PROGRAM PRG_Seq
VAR
    eStep, ePrevStep : E_Step := E_Step.eInit;
    nFaultCode       : UINT;        // 1=E-stop 2=no air 3=cylinder fault 4=step timeout
    nPartCount       : UDINT;
    bRejectPart      : BOOL;
    xAutoRun         : BOOL;
    xReady           : BOOL;
    xEnableCyl       : BOOL;

    // cylinder commands (TRUE = working position AS, FALSE = home GS) - persistent
    xInfeedWork, xClampWork, xEjectWork, xDivertWork, xOutfeedWork : BOOL;
    // momentary commands (cleared every scan, set by the active step)
    xBlow, xBypass, xLaserOn, xTrig : BOOL;

    fbInfeed, fbOutfeed, fbEjector, fbClamp, fbDiverter : FB_Cylinder;
    rStart, rReset   : R_TRIG;
    fbPart           : TON;
    fbBlowTime       : TON;
    fbStepTO         : TON;
    tStepTimeout     : TIME := T#30S;
    tBlow            : TIME := T#1S;
    tPartDebounce    : TIME := T#200MS;
END_VAR

rStart(CLK := GVL_Ctrl.xStart);
rReset(CLK := GVL_Ctrl.xReset);
IF rStart.Q THEN xAutoRun := TRUE;  END_IF
IF GVL_Ctrl.xStop THEN xAutoRun := FALSE; END_IF

// momentary outputs default to OFF every scan
xBlow := FALSE;  xBypass := FALSE;  xLaserOn := FALSE;  xTrig := FALSE;

xReady := GVL_IO.xPressureOK AND NOT GVL_IO.xEStop
          AND GVL_IO.xServoInLatched AND GVL_IO.xServoOutLatched;
xEnableCyl := (eStep <> E_Step.eFault) AND NOT GVL_IO.xEStop AND GVL_IO.xPressureOK;

// ---- cylinders (called first so that feedback is current for the transitions)
fbInfeed(  xCmdWork := xInfeedWork,  xEnable := xEnableCyl, xReset := rReset.Q,
           xSensWork := GVL_IO.stInfeed.xSensWork,   xSensHome := GVL_IO.stInfeed.xSensHome,
           xValveWork => GVL_IO.stInfeed.xValveWork, xValveHome => GVL_IO.stInfeed.xValveHome);
fbOutfeed( xCmdWork := xOutfeedWork, xEnable := xEnableCyl, xReset := rReset.Q,
           xSensWork := GVL_IO.stOutfeed.xSensWork,   xSensHome := GVL_IO.stOutfeed.xSensHome,
           xValveWork => GVL_IO.stOutfeed.xValveWork, xValveHome => GVL_IO.stOutfeed.xValveHome);
fbEjector( xCmdWork := xEjectWork,   xEnable := xEnableCyl, xReset := rReset.Q,
           xSensWork := GVL_IO.stEjector.xSensWork,   xSensHome := GVL_IO.stEjector.xSensHome,
           xValveWork => GVL_IO.stEjector.xValveWork, xValveHome => GVL_IO.stEjector.xValveHome);
fbClamp(   xCmdWork := xClampWork,   xEnable := xEnableCyl, xReset := rReset.Q,
           xSensWork := GVL_IO.stClamp.xSensWork,   xSensHome := GVL_IO.stClamp.xSensHome,
           xValveWork => GVL_IO.stClamp.xValveWork, xValveHome => GVL_IO.stClamp.xValveHome);
fbDiverter(xCmdWork := xDivertWork,  xEnable := xEnableCyl, xReset := rReset.Q,
           xSensWork := GVL_IO.stDiverter.xSensWork,   xSensHome := GVL_IO.stDiverter.xSensHome,
           xValveWork => GVL_IO.stDiverter.xValveWork, xValveHome => GVL_IO.stDiverter.xValveHome);

// ---- step timeout (restarts whenever the step changes)
fbStepTO(IN := (eStep = ePrevStep) AND (eStep <> E_Step.eIdle) AND (eStep <> E_Step.eWaitPart)
               AND (eStep <> E_Step.eFault),
         PT := tStepTimeout);
ePrevStep := eStep;

// ---- supervision
IF eStep <> E_Step.eFault THEN
    IF GVL_IO.xEStop THEN
        nFaultCode := 1;  eStep := E_Step.eFault;
    ELSIF NOT GVL_IO.xPressureOK THEN
        nFaultCode := 2;  eStep := E_Step.eFault;
    ELSIF fbInfeed.xFault OR fbOutfeed.xFault OR fbEjector.xFault OR fbClamp.xFault OR fbDiverter.xFault THEN
        nFaultCode := 3;  eStep := E_Step.eFault;
    ELSIF fbStepTO.Q THEN
        nFaultCode := 4;  eStep := E_Step.eFault;
    END_IF
END_IF

// ---- sequence
fbPart(IN := GVL_IO.xLS_Infeed, PT := tPartDebounce);
fbBlowTime(IN := (eStep = E_Step.eBlowOff), PT := tBlow);

CASE eStep OF

    E_Step.eInit:
        xInfeedWork := FALSE;  xClampWork := FALSE;  xEjectWork := FALSE;
        xDivertWork := FALSE;  xOutfeedWork := FALSE;
        IF fbInfeed.xInHome AND fbOutfeed.xInHome AND fbEjector.xInHome
           AND fbClamp.xInHome AND fbDiverter.xInHome THEN
            eStep := E_Step.eIdle;
        END_IF

    E_Step.eIdle:
        IF xAutoRun AND xReady THEN
            eStep := E_Step.eWaitPart;
        END_IF

    E_Step.eWaitPart:
        IF NOT xAutoRun THEN
            eStep := E_Step.eIdle;
        ELSIF fbPart.Q THEN
            bRejectPart := GVL_Ctrl.xReject;      // latch quality decision for this part
            eStep := E_Step.eInfeedFwd;
        END_IF

    E_Step.eInfeedFwd:
        xInfeedWork := TRUE;
        IF fbInfeed.xInWork THEN eStep := E_Step.eClampFwd; END_IF

    E_Step.eClampFwd:
        xClampWork := TRUE;
        IF fbClamp.xInWork THEN eStep := E_Step.eInfeedBack; END_IF

    E_Step.eInfeedBack:
        xInfeedWork := FALSE;
        IF fbInfeed.xInHome THEN eStep := E_Step.eLoadJob; END_IF

    E_Step.eLoadJob:
        xLaserOn := TRUE;                          // LaserEnable + STO release + job select
        IF GVL_IO.xCW_JobLoaded AND GVL_IO.xCW_Lready THEN
            eStep := E_Step.eLaserRun;
        END_IF

    E_Step.eLaserRun:
        xLaserOn := TRUE;  xTrig := TRUE;
        IF GVL_IO.xCW_MarkBusy THEN eStep := E_Step.eLaserWait; END_IF

    E_Step.eLaserWait:
        xLaserOn := TRUE;  xTrig := TRUE;
        IF NOT GVL_IO.xCW_MarkBusy THEN eStep := E_Step.eBlowOff; END_IF

    E_Step.eBlowOff:
        xBlow := TRUE;
        IF fbBlowTime.Q THEN eStep := E_Step.eClampBack; END_IF

    E_Step.eClampBack:
        xClampWork := FALSE;
        IF fbClamp.xInHome THEN eStep := E_Step.eDiverter; END_IF

    E_Step.eDiverter:
        xDivertWork := bRejectPart;                // work = reject path, home = good path
        IF (bRejectPart AND fbDiverter.xInWork) OR (NOT bRejectPart AND fbDiverter.xInHome) THEN
            eStep := E_Step.eEject;
        END_IF

    E_Step.eEject:
        xEjectWork := TRUE;
        xBypass := bRejectPart;                    // bypass valve only for rejects
        IF fbEjector.xInWork THEN eStep := E_Step.eEjectBack; END_IF

    E_Step.eEjectBack:
        xEjectWork := FALSE;
        xBypass := bRejectPart;
        IF fbEjector.xInHome THEN
            IF bRejectPart THEN
                eStep := E_Step.eCycleEnd;         // reject left through bypass
            ELSE
                eStep := E_Step.eOutfeedWait;
            END_IF
        END_IF

    E_Step.eOutfeedWait:
        IF GVL_IO.xLS_Outfeed THEN eStep := E_Step.eOutfeed; END_IF

    E_Step.eOutfeed:
        xOutfeedWork := TRUE;
        IF fbOutfeed.xInWork THEN eStep := E_Step.eOutfeedBack; END_IF

    E_Step.eOutfeedBack:
        xOutfeedWork := FALSE;
        IF fbOutfeed.xInHome THEN eStep := E_Step.eCycleEnd; END_IF

    E_Step.eCycleEnd:
        xDivertWork := FALSE;
        IF fbDiverter.xInHome THEN
            nPartCount := nPartCount + 1;
            eStep := E_Step.eIdle;
        END_IF

    E_Step.eFault:
        xAutoRun := FALSE;
        IF rReset.Q AND NOT GVL_IO.xEStop AND GVL_IO.xPressureOK THEN
            nFaultCode := 0;
            eStep := E_Step.eInit;
        END_IF

END_CASE

// ---- write logic outputs
GVL_IO.xVent        := GVL_IO.xEStop;                       // vent maintenance unit on E-stop
GVL_IO.xLaserEnable := xLaserOn AND xEnableCyl;
GVL_IO.xCW_STO      := xLaserOn AND xEnableCyl;             // ASSUMPTION: TRUE = STO released
GVL_IO.xCW_Trig     := xTrig    AND xEnableCyl;
IF xLaserOn THEN GVL_IO.nCW_Job := GVL_Ctrl.nJobNo; ELSE GVL_IO.nCW_Job := 0; END_IF
GVL_IO.xBlowAS      := xBlow   AND xEnableCyl;
GVL_IO.xBlowGS      := xEnableCyl AND NOT xBlow;
GVL_IO.xBypassAS    := xBypass AND xEnableCyl;
GVL_IO.xBypassGS    := xEnableCyl AND NOT xBypass;

END_PROGRAM

(* stored: Version 1.1.0.1
   POU PRG_Seq: Id {7da9cb7f-2a2b-433f-a108-ae73eb091758}, SpecialFunc None *)
